// TIA Portal V18 export
TYPE "Config_SEND_RCV"
   STRUCT
      modezone { S7_SetPoint := 'True'} : Array[1.."ModeZone_Setup_Const"] of "Comm";
   END_STRUCT;
END_TYPE
